Universal Robots URScript: T008_zai-org_GLM-4.7-FP8_edit_perf_rep1.urscript

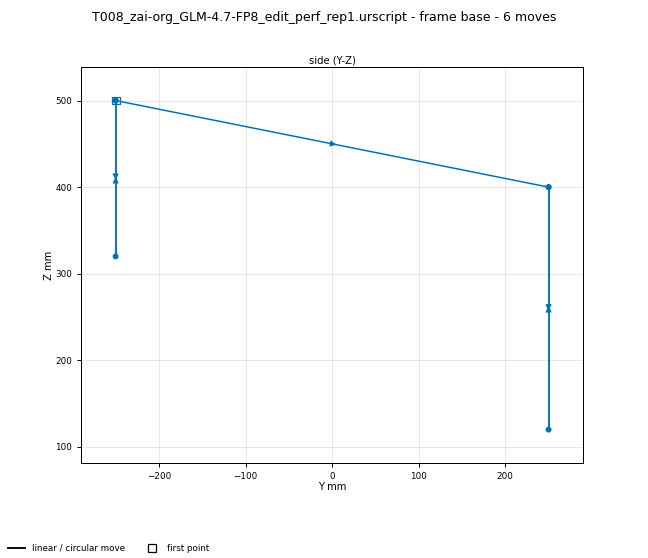
[picture p0: tool path of T008_zai-org_GLM-4.7-FP8_edit_perf_rep1.urscript in frame base, 6 of 8 moves have a stored position in this frame; points joined in program order, loops and branches not executed]
# Task: T008 — Heavy depalletizing — fenced mode (Optimized)
# Generated by ENFIELD IR→URScript Translator
# Operating mode: fenced | Max TCP speed: 0.450 m/s
# Robot: ur5e
#
# WARNING: This is auto-generated code for SIMULATION ONLY.
# Do NOT deploy to a physical robot without safety review.

def task_T008():
  # [0] Verify E-Stop
  # E-Stop safety check (hardware-enforced on UR controller)
  if (get_digital_in(0) == True):
    popup("E-Stop active — aborting program.", error=True)
    halt
  end

  # [1] Home
  # Optimized: Increased joint velocity and acceleration for faster transit
  movej([0.0000, -1.5708, 1.5708, -1.5708, -1.5708, 0.0000], a=2.5000, v=1.8000)

  # [2] Above pallet
  # Optimized: Increased velocity to max TCP limit (0.45 m/s), increased blend radius
  movel(p[0.500000, -0.250000, 0.500000, 0.0000, 3.1416, 0.0000], a=1.5000, v=0.4500, r=0.0500)

  # [3] Descend to top layer
  # Optimized: Increased approach speed for faster cycle time
  movel(p[0.500000, -0.250000, 0.320000, 0.0000, 3.1416, 0.0000], a=1.0000, v=0.3000)

  # [4] Gripper CLOSE
  # Gripper CLOSE (force=120 N)
  set_digital_out(0, True)

  # [5] Grip settle
  # Optimized: Reduced sleep time to minimum required for gripper actuation
  sleep(0.2000)

  # [6] Lift box
  # Optimized: Increased lift speed and blend radius for smoother transition
  movel(p[0.500000, -0.250000, 0.500000, 0.0000, 3.1416, 0.0000], a=1.2000, v=0.3500, r=0.0500)

  # [7] Transit to conveyor
  # Optimized: Increased velocity to max TCP limit, increased blend radius
  movel(p[0.500000, 0.250000, 0.400000, 0.0000, 3.1416, 0.0000], a=1.5000, v=0.4500, r=0.0500)

  # [8] Place on conveyor
  # Optimized: Increased placement speed
  movel(p[0.500000, 0.250000, 0.120000, 0.0000, 3.1416, 0.0000], a=1.0000, v=0.2500)

  # [9] Gripper OPEN
  # Gripper OPEN
  set_digital_out(0, False)

  # [10] Release settle
  # Optimized: Reduced sleep time
  sleep(0.1000)

  # [11] Retract
  # Optimized: Increased velocity to max TCP limit, increased blend radius
  movel(p[0.500000, 0.250000, 0.400000, 0.0000, 3.1416, 0.0000], a=1.5000, v=0.4500, r=0.0500)

  # [12] Return home
  # Optimized: Increased joint velocity and acceleration
  movej([0.0000, -1.5708, 1.5708, -1.5708, -1.5708, 0.0000], a=2.5000, v=1.8000)

end

# Entry point
task_T008()
